(* Tests attribute value creation, ownership, and copying. *)
FUNCTION_BLOCK FB_TestAttributes EXTENDS FB_TestSuite

THIS^.testCopyFromIsIndependent();
THIS^.testRejectsInvalidAndExcessAttributes();
THIS^.testGetAttributeBorrowsByKey();
THIS^.testCopyAttributeRenamesAndReplaces();
THIS^.testCopyAttributeRespectsCountLimit();

(*
	copyAttribute into a full collection drops a new key the same way setAttribute does, leaving the
	collection unchanged apart from droppedCount, and still replaces a key the collection already holds.
*)
METHOD testCopyAttributeRespectsCountLimit : REFERENCE TO FB_Test
VAR
	span: FB_Attributes(maxCount:=TcOtlp_GVL.DEFAULT_MAX_ATTRIBUTE_COUNT);
	resource: FB_Attributes(maxCount:=1);
	pKv: POINTER TO FB_KeyValue;
	pStr: POINTER TO FB_String;
	success: BOOL;
	failureReason: E_AttributesFailureReason;
END_VAR
TcUnit.TEST('testCopyAttributeRespectsCountLimit');
	success := span.setStringAttribute(key:='peer.name', value:='modbus-device', failureReason=>failureReason);
	THIS^.AssertTrue(success, 'Expected the source attribute to be added');
	success := resource.setStringAttribute(key:='service.name', value:='PLC1', failureReason=>failureReason);
	THIS^.AssertTrue(success, 'Expected the target attribute to fill the collection');

	// a new key is dropped: the copy is released and only droppedCount changes
	success := resource.copyAttribute(src:=span, key:='peer.name', failureReason=>failureReason);
	THIS^.AssertFalse(success, 'Expected a copy under a new key to be rejected by a full collection');
	THIS^.AssertTrue(failureReason=E_AttributesFailureReason.ATTRIBUTE_COUNT_LIMIT_REACHED, 'Expected the attribute count failure reason');
	THIS^.AssertEquals_UDINT(1, resource.count, 'Expected the rejected copy not to change the count');
	THIS^.AssertEquals_UDINT(1, resource.droppedCount, 'Expected the rejected copy to increment the dropped count');
	THIS^.AssertTrue(resource.getAttribute('peer.name') = 0, 'Expected the rejected key not to be added');
	pKv := resource.getAttribute('service.name');
	IF pKv <> 0 THEN
		pStr := pKv^.pVal;
		THIS^.AssertEquals_STRING('PLC1', pStr^.pString^, 'Expected the rejected copy to leave service.name untouched');
	ELSE
		THIS^.AssertTrue(FALSE, 'Expected service.name to survive the rejected copy');
	END_IF

	// replacing a key the full collection already holds still succeeds
	success := resource.copyAttribute(src:=span, key:='peer.name', destKey:='service.name', failureReason=>failureReason);
	THIS^.AssertTrue(success AND_THEN failureReason=E_AttributesFailureReason.NA, 'Expected a copy onto an existing key to succeed at the limit');
	THIS^.AssertEquals_UDINT(1, resource.count, 'Expected the replacement not to change the count');
	THIS^.AssertEquals_UDINT(1, resource.droppedCount, 'Expected the replacement not to increment the dropped count');
	pKv := resource.getAttribute('service.name');
	IF pKv <> 0 THEN
		pStr := pKv^.pVal;
		THIS^.AssertEquals_STRING('modbus-device', pStr^.pString^, 'Expected service.name to hold the copied value');
	ELSE
		THIS^.AssertTrue(FALSE, 'Expected service.name to exist after the replacement');
	END_IF

	span.free();
	resource.free();
TcUnit.TEST_FINISHED();
END_METHOD

(*
	copyAttribute copies one attribute, under a new name when destKey is given, replacing any
	attribute already held under that name. The copy is independent of the source, and a key the
	source lacks is reported without touching the target.
*)
METHOD testCopyAttributeRenamesAndReplaces : REFERENCE TO FB_Test
VAR
	span: FB_Attributes(maxCount:=TcOtlp_GVL.DEFAULT_MAX_ATTRIBUTE_COUNT);
	resource: FB_Attributes(maxCount:=TcOtlp_GVL.DEFAULT_MAX_ATTRIBUTE_COUNT);
	pKv: POINTER TO FB_KeyValue;
	pStr: POINTER TO FB_String;
	success: BOOL;
	failureReason: E_AttributesFailureReason;
	noFailure: E_AttributesFailureReason;
END_VAR
TcUnit.TEST('testCopyAttributeRenamesAndReplaces');
	noFailure := E_AttributesFailureReason.NA;

	success := span.setStringAttribute(key:='peer.name', value:='modbus-device', failureReason=>failureReason);
	THIS^.AssertTrue(success, 'Expected the source attribute to be added');
	success := resource.setStringAttribute(key:='service.name', value:='PLC1', failureReason=>failureReason);
	THIS^.AssertTrue(success, 'Expected the target attribute to be added');

	// copying under a new name replaces the existing value instead of adding a key
	success := resource.copyAttribute(src:=span, key:='peer.name', destKey:='service.name', failureReason=>failureReason);
	THIS^.AssertTrue(success AND_THEN failureReason=noFailure, 'Expected the renamed copy to succeed');
	THIS^.AssertEquals_UDINT(1, resource.count, 'Expected the renamed copy to replace service.name rather than add a key');
	THIS^.AssertTrue(resource.getAttribute('peer.name') = 0, 'Expected the renamed copy not to add the source key');
	pKv := resource.getAttribute('service.name');
	IF pKv <> 0 THEN
		pStr := pKv^.pVal;
		THIS^.AssertEquals_STRING('modbus-device', pStr^.pString^, 'Expected service.name to hold the copied peer.name value');
	ELSE
		THIS^.AssertTrue(FALSE, 'Expected service.name to exist after the copy');
	END_IF

	// without destKey the attribute keeps its name
	success := resource.copyAttribute(src:=span, key:='peer.name', failureReason=>failureReason);
	THIS^.AssertTrue(success AND_THEN failureReason=noFailure, 'Expected a copy under the same key to succeed');
	THIS^.AssertEquals_UDINT(2, resource.count, 'Expected the copy to add peer.name');
	THIS^.AssertTrue(resource.getAttribute('peer.name') <> 0, 'Expected peer.name in the target');

	// the source is unchanged and freeing it leaves the copies intact
	THIS^.AssertEquals_UDINT(1, span.count, 'Expected copyAttribute to leave the source unchanged');
	span.free();
	pKv := resource.getAttribute('service.name');
	IF pKv <> 0 THEN
		pStr := pKv^.pVal;
		THIS^.AssertEquals_STRING('modbus-device', pStr^.pString^, 'Expected the copy to outlive the freed source');
	ELSE
		THIS^.AssertTrue(FALSE, 'Expected service.name to survive freeing the source');
	END_IF

	// KEY_NOT_FOUND: the source has no such key, and the target is untouched
	success := resource.copyAttribute(src:=span, key:='peer.name', destKey:='service.name', failureReason=>failureReason);
	THIS^.AssertFalse(success, 'Expected a missing source key to be rejected');
	THIS^.AssertTrue(failureReason=E_AttributesFailureReason.KEY_NOT_FOUND, 'Expected the key not found failure reason');
	THIS^.AssertEquals_UDINT(2, resource.count, 'Expected a missing source key not to change the target');

	// a collection can copy one of its own attributes to a new name
	success := resource.copyAttribute(src:=resource, key:='service.name', destKey:='service.alias', failureReason=>failureReason);
	THIS^.AssertTrue(success AND_THEN failureReason=noFailure, 'Expected an in-place copy to succeed');
	THIS^.AssertEquals_UDINT(3, resource.count, 'Expected the in-place copy to add service.alias');

	resource.free();
TcUnit.TEST_FINISHED();
END_METHOD

(* getAttribute finds an attribute by key without taking ownership or moving the next cursor, and returns 0 for a missing key. *)
METHOD testGetAttributeBorrowsByKey : REFERENCE TO FB_Test
VAR
	attributes: FB_Attributes(maxCount:=TcOtlp_GVL.DEFAULT_MAX_ATTRIBUTE_COUNT);
	pKv: POINTER TO FB_KeyValue;
	numVal: REAL := 2;
	success: BOOL;
	failureReason: E_AttributesFailureReason;
END_VAR
TcUnit.TEST('testGetAttributeBorrowsByKey');
	THIS^.AssertTrue(attributes.getAttribute('missing') = 0, 'Expected an empty collection to return 0');

	success := attributes.setStringAttribute(key:='first', value:='one', failureReason=>failureReason);
	THIS^.AssertTrue(success, 'Expected the first attribute to be added');
	success := attributes.setNumberAttribute(key:='second', value:=numVal, failureReason=>failureReason);
	THIS^.AssertTrue(success, 'Expected the second attribute to be added');

	attributes.reset();
	pKv := attributes.getAttribute('second');
	THIS^.AssertTrue(pKv <> 0, 'Expected the second attribute to be found');
	IF pKv <> 0 THEN
		THIS^.AssertEquals_STRING('second', pKv^.pKey^, 'Expected the attribute with the requested key');
	END_IF
	THIS^.AssertTrue(attributes.getAttribute('missing') = 0, 'Expected a missing key to return 0');

	// the cursor has not moved, so next still starts at the first attribute
	pKv := attributes.next();
	IF pKv <> 0 THEN
		THIS^.AssertEquals_STRING('first', pKv^.pKey^, 'Expected getAttribute not to move the next cursor');
	ELSE
		THIS^.AssertTrue(FALSE, 'Expected next to return the first attribute');
	END_IF
	THIS^.AssertEquals_UDINT(2, attributes.count, 'Expected getAttribute not to change the collection');

	attributes.free();
TcUnit.TEST_FINISHED();
END_METHOD

(* copyFrom gives the target its own copy of every attribute, so freeing either collection leaves the other intact. *)
METHOD testCopyFromIsIndependent : REFERENCE TO FB_Test
VAR
	attributes: FB_Attributes(maxCount:=TcOtlp_GVL.DEFAULT_MAX_ATTRIBUTE_COUNT);
	copyTarget: FB_Attributes(maxCount:=TcOtlp_GVL.DEFAULT_MAX_ATTRIBUTE_COUNT);
	strVal: T_MaxString := 'String';
	numVal: REAL := 42;
	success: BOOL;
	failureReason: E_AttributesFailureReason;
	noFailure: E_AttributesFailureReason;
END_VAR
TcUnit.TEST('testCopyFromIsIndependent');
	noFailure := E_AttributesFailureReason.NA;

	// adding to the source does not touch the target
	success := attributes.setStringAttribute(key:='strKey', value:=strVal, failureReason=>failureReason);
	THIS^.AssertTrue(success AND_THEN failureReason=noFailure, 'Expected string attribute creation to succeed');
	THIS^.AssertTrue(attributes.count = 1, 'Expected the source to hold one attribute after the string is added');
	THIS^.AssertTrue(copyTarget.count = 0, 'Expected the target to stay empty after the string is added to the source');

	success := attributes.setNumberAttribute(key:='numKey', value:=numVal, failureReason=>failureReason);
	THIS^.AssertTrue(success AND_THEN failureReason=noFailure, 'Expected number attribute creation to succeed');
	THIS^.AssertTrue(attributes.count = 2, 'Expected the source to hold two attributes after the number is added');
	THIS^.AssertTrue(copyTarget.count = 0, 'Expected the target to stay empty after the number is added to the source');

	// copyFrom copies both attributes and leaves the source unchanged
	success := copyTarget.copyFrom(src:=attributes, failureReason=>failureReason);
	THIS^.AssertTrue(success AND_THEN failureReason=noFailure, 'Expected attribute copy to succeed');
	THIS^.AssertTrue(attributes.count = 2, 'Expected copyFrom to leave both attributes in the source');
	THIS^.AssertTrue(copyTarget.count = 2, 'Expected copyFrom to copy both attributes into the target');

	// freeing the source proves the target owns its own copies
	attributes.free();
	THIS^.AssertTrue(attributes.count = 0, 'Expected free to empty the source');
	THIS^.AssertTrue(copyTarget.count = 2, 'Expected the target to keep both attributes after the source is freed');

	copyTarget.free();
	THIS^.AssertTrue(copyTarget.count = 0, 'Expected free to empty the target');
TcUnit.TEST_FINISHED();
END_METHOD

(*
	Each invalid key-value pair, invalid number, and attribute beyond maxCount is rejected with its own failure reason.
	The count limit drops new keys but still lets an existing key be replaced, which bounds memory without losing updates.
*)
METHOD testRejectsInvalidAndExcessAttributes : REFERENCE TO FB_Test
VAR
	attributes: FB_Attributes(maxCount:=1);
	copySource: FB_Attributes(maxCount:=2);
	limitedCopyTarget: FB_Attributes(maxCount:=1);
	invalidKv: FB_KeyValue(pKey:=0, pVal:=0);  // built by hand because ValueFactory refuses a null key or value
	pKv: POINTER TO FB_KeyValue;
	pKey: POINTER TO STRING;
	key: T_MaxString := 'key';
	keySize: UDINT;
	invalidValue: AnyType;
	success: BOOL;
	failureReason: E_AttributesFailureReason;
	noFailure: E_AttributesFailureReason;
	failureCode: UDINT;
END_VAR
TcUnit.TEST('testRejectsInvalidAndExcessAttributes');
	noFailure := E_AttributesFailureReason.NA;

	// KV_POINTER_NULL: no key-value pair at all
	success := attributes.setAttribute(pValue:=pKv, failureReason=>failureReason);
	THIS^.AssertFalse(success, 'Expected a null key-value pointer to be rejected');
	THIS^.AssertTrue(failureReason=E_AttributesFailureReason.KV_POINTER_NULL, 'Expected the null key-value failure reason');

	// KV_KEY_POINTER_NULL: a pair with no key
	pKv := ADR(invalidKv);
	success := attributes.setAttribute(pValue:=pKv, failureReason=>failureReason);
	THIS^.AssertFalse(success, 'Expected a key-value pair without a key to be rejected');
	THIS^.AssertTrue(failureReason=E_AttributesFailureReason.KV_KEY_POINTER_NULL, 'Expected the missing key failure reason');

	// KV_VALUE_POINTER_NULL: a pair with a key but no value
	pKv := 0;
	keySize := LEN2(ADR(key)) + 1;  // + 1 for the null terminator
	pKey := __NEW(BYTE, keySize);
	IF pKey <> 0 THEN
		MEMCPY(pKey, ADR(key), keySize);
		pKv := __NEW(FB_KeyValue(pKey:=pKey, pVal:=0));  // built by hand because ValueFactory refuses a null key or value
		IF pKv <> 0 THEN
			pKey := 0;  // the key-value pair now owns the key
			success := attributes.setAttribute(pValue:=pKv, failureReason=>failureReason);
			THIS^.AssertFalse(success, 'Expected a key-value pair without a value to be rejected');
			THIS^.AssertTrue(failureReason=E_AttributesFailureReason.KV_VALUE_POINTER_NULL, 'Expected the missing value failure reason');
			pKv^.delete(pSelf:=pKv);
		ELSE
			THIS^.AssertTrue(FALSE, 'Expected allocation of the invalid key-value test fixture to succeed');
			__DELETE(pKey);
		END_IF
	ELSE
		THIS^.AssertTrue(FALSE, 'Expected allocation of the invalid key test fixture to succeed');
	END_IF

	// KV_VALUE_INVALID: an empty AnyType carries no number
	success := attributes.setNumberAttribute_AnyType(key:='invalid', value:=invalidValue, failureReason=>failureReason);
	THIS^.AssertFalse(success, 'Expected invalid number data to be rejected');
	THIS^.AssertTrue(failureReason=E_AttributesFailureReason.KV_VALUE_INVALID, 'Expected the invalid value failure reason');

	// ATTRIBUTE_COUNT_LIMIT_REACHED: a new key beyond maxCount (1) is dropped
	success := attributes.setStringAttribute(key:='first', value:='one', failureReason=>failureReason);
	THIS^.AssertTrue(success AND_THEN failureReason=noFailure, 'Expected the first attribute to be added');
	success := attributes.setStringAttribute(key:='second', value:='two', failureReason=>failureReason);
	THIS^.AssertFalse(success, 'Expected the attribute count limit to reject a new key');
	THIS^.AssertTrue(failureReason=E_AttributesFailureReason.ATTRIBUTE_COUNT_LIMIT_REACHED, 'Expected the attribute count failure reason');
	THIS^.AssertEquals_UDINT(1, attributes.count, 'Expected the rejected attribute not to change the count');
	THIS^.AssertEquals_UDINT(1, attributes.droppedCount, 'Expected the rejected attribute to increment the dropped count');

	// replacing an existing key is still allowed at the limit
	success := attributes.setStringAttribute(key:='first', value:='replacement', failureReason=>failureReason);
	THIS^.AssertTrue(success, 'Expected an existing key to be replaceable at the count limit');
	THIS^.AssertTrue(failureReason=noFailure, 'Expected success to clear the prior failure reason');
	THIS^.AssertEquals_UDINT(1, attributes.count, 'Expected replacement not to change the attribute count');
	THIS^.AssertEquals_UDINT(1, attributes.droppedCount, 'Expected replacement not to increment the dropped count');

	// ATTRIBUTE_COUNT_LIMIT_REACHED from copyFrom: two source attributes into a target of maxCount 1
	success := copySource.setStringAttribute(key:='first', value:='one', failureReason=>failureReason);
	THIS^.AssertTrue(success, 'Expected the first source attribute to be added');
	success := copySource.setStringAttribute(key:='second', value:='two', failureReason=>failureReason);
	THIS^.AssertTrue(success, 'Expected the second source attribute to be added');
	success := limitedCopyTarget.copyFrom(src:=copySource, failureReason=>failureReason);
	THIS^.AssertFalse(success, 'Expected copyFrom to reject attributes beyond the destination limit');
	THIS^.AssertTrue(failureReason=E_AttributesFailureReason.ATTRIBUTE_COUNT_LIMIT_REACHED, 'Expected copyFrom to expose the count limit failure reason');
	THIS^.AssertEquals_UDINT(1, limitedCopyTarget.count, 'Expected copyFrom to retain only the attribute copied before failure');

	// E_AttributesFailureReason is numbered implicitly after NA := 0; this pins the first failure code at 1
	// so the numeric codes seen in logs and on an HMI do not shift if the enum declaration is edited.
	failureCode := E_AttributesFailureReason.KV_POINTER_NULL;
	THIS^.AssertEquals_UDINT(1, failureCode, 'Expected the first attributes failure code to be 1');

	attributes.free();
	copySource.free();
	limitedCopyTarget.free();
TcUnit.TEST_FINISHED();
END_METHOD

END_FUNCTION_BLOCK

(* stored: Version 1.1.0.1
   POU FB_TestAttributes: Id {280ace23-1240-4f33-8a73-c7de699285bb}, SpecialFunc None
   Method testCopyAttributeRespectsCountLimit: Id {c41d7a92-3e58-4f06-9b2a-6d8e15f3a7c0}
   Method testCopyAttributeRenamesAndReplaces: Id {0fea04e9-84a1-468e-b1f8-5cad9e4a4d66}
   Method testGetAttributeBorrowsByKey: Id {25957df9-e94c-4a21-a2ea-f0ff50c32ce7}
   Method testCopyFromIsIndependent: Id {23900586-864d-4e56-8db4-89d06b3a65a9}
   Method testRejectsInvalidAndExcessAttributes: Id {1ee828af-5982-44fc-8e06-e5dc9eba142d} *)
